                            IF #statSendBufferPos + #tempBytesUsedUtf8 <=  THEN
                              #statUserNamePos += 1;
                              CASE #tempBytesUsedUtf8 OF
                                :  // Statement section case 1
                                  #statSendBuffer[#statSendBufferPos] := #tempConvertedUtf8.%B0;
                                  #statSendBufferPos += 1;
                                :
                                  #statSendBuffer[#statSendBufferPos] := #tempConvertedUtf8.%B0;
                                  #statSendBufferPos += 1;
                                  #statSendBuffer[#statSendBufferPos] := #tempConvertedUtf8.%B1;
                                  #statSendBufferPos += 1;
                                :  // Statement section case 2 to 4
                                  #statSendBuffer[#statSendBufferPos] := #tempConvertedUtf8.%B0;
                                  #statSendBufferPos += 1;
                                  #statSendBuffer[#statSendBufferPos] := #tempConvertedUtf8.%B1;
                                  #statSendBufferPos += 1;
                                  #statSendBuffer[#statSendBufferPos] := #tempConvertedUtf8.%B2;
                                  #statSendBufferPos += 1;
                                ELSE  // Statement section ELSE
                                  ;
                              END_CASE;
                            ELSE
                              //When buffer full
                              EXIT;
                            END_IF;
                          END_FOR;
                          IF #statUserNamePos >= LEN(#username) THEN
                            #statUserNameEncodeState := ;
                          END_IF;

                        ELSE  // Statement section ELSE
                          ;
                      END_CASE;
                    END_IF;

                    // Password
                    // If the Password Flag is set to 1, the Password the next field in the payload. It must be > 0 Bytes
                    //Password field contains 0 to 65535 bytes OF binary data prefixed with a two Byte length field which indicates the number OF bytes used

                    IF #statClientIdEncodeState =
                      AND (#statWillTopicEncodeState =  OR #statWillTopicEncodeState = )
                      AND (#statWillMessageEncodeState =  OR #statWillMessageEncodeState = )
                      AND (#statUserNameEncodeState =  OR #statUserNameEncodeState = )
                      AND #statSendBufferPos <=  -  THEN
                      //When Will Topic and Will Message is encoded and buffer not full
                      CASE #statPasswordEncodeState OF
                        :  // Statement section case 1
                          //ADD len info into paket

                          #tempWordForSliceAddress := UINT_TO_WORD(#statPasswordLenUtf8Encoded);
                          #statSendBuffer[#statSendBufferPos] := #tempWordForSliceAddress.%B1; //MSB
                          #statSendBufferPos += 1;
                          #statSendBuffer[#statSendBufferPos] := #tempWordForSliceAddress.%B0; // LSB
                          #statSendBufferPos += 1;

                          FOR #tempLoopCounter := #statPasswordPos TO LEN(#password) DO
                            LMQTT_ConvertToUtf8(character     := #password[#tempLoopCounter],
                                                  convertedUtf8 => #tempConvertedUtf8,
                                                  bytesUsed     => #tempBytesUsedUtf8,
                                                  error         => #tempErrorConvertUtf8,
                                                  status        => #tempStatusConvertUtf8);

                            IF #statSendBufferPos + #tempBytesUsedUtf8 <=  THEN
                              //Increment when successful
                              #statPasswordPos += 1;

                              CASE #tempBytesUsedUtf8 OF
                                :  // Statement section case 1
                                  #statSendBuffer[#statSendBufferPos] := #tempConvertedUtf8.%B0;
                                  #statSendBufferPos += 1;
                                :
                                  #statSendBuffer[#statSendBufferPos] := #tempConvertedUtf8.%B0;
                                  #statSendBufferPos += 1;
                                  #statSendBuffer[#statSendBufferPos] := #tempConvertedUtf8.%B1;
                                  #statSendBufferPos += 1;
                                :  // Statement section case 2 to 4
                                  #statSendBuffer[#statSendBufferPos] := #tempConvertedUtf8.%B0;
                                  #statSendBufferPos += 1;
                                  #statSendBuffer[#statSendBufferPos] := #tempConvertedUtf8.%B1;
                                  #statSendBufferPos += 1;
                                  #statSendBuffer[#statSendBufferPos] := #tempConvertedUtf8.%B2;
                                  #statSendBufferPos += 1;
                                ELSE  // Statement section ELSE
                                  ;
                              END_CASE;
                            ELSE
                              //When buffer full
                              #statPasswordEncodeState := ;
                              EXIT;
                            END_IF;
                          END_FOR;

                          IF #statPasswordPos >= LEN(#password) THEN
                            #statPasswordEncodeState := ;
                          END_IF;

                        :  // Statement section case 2 to 4
                          FOR #tempLoopCounter := #statPasswordPos TO LEN(#password) DO
                            LMQTT_ConvertToUtf8(character     := #password[#tempLoopCounter],
                                                  convertedUtf8 => #tempConvertedUtf8,
                                                  bytesUsed     => #tempBytesUsedUtf8,
                                                  error         => #tempErrorConvertUtf8,
                                                  status        => #tempStatusConvertUtf8);

                            IF #statSendBufferPos + #tempBytesUsedUtf8 <=  THEN
                              #statPasswordPos += 1;
                              CASE #tempBytesUsedUtf8 OF
                                :  // Statement section case 1
                                  #statSendBuffer[#statSendBufferPos] := #tempConvertedUtf8.%B0;
                                  #statSendBufferPos += 1;
                                :
                                  #statSendBuffer[#statSendBufferPos] := #tempConvertedUtf8.%B0;
                                  #statSendBufferPos += 1;
                                  #statSendBuffer[#statSendBufferPos] := #tempConvertedUtf8.%B1;
                                  #statSendBufferPos += 1;
                                :  // Statement section case 2 to 4
                                  #statSendBuffer[#statSendBufferPos] := #tempConvertedUtf8.%B0;
                                  #statSendBufferPos += 1;
                                  #statSendBuffer[#statSendBufferPos] := #tempConvertedUtf8.%B1;
                                  #statSendBufferPos += 1;
                                  #statSendBuffer[#statSendBufferPos] := #tempConvertedUtf8.%B2;
                                  #statSendBufferPos += 1;
                                ELSE  // Statement section ELSE
                                  ;
                              END_CASE;
                            ELSE
                              //When buffer full
                              EXIT;
                            END_IF;
                          END_FOR;
                          IF #statPasswordPos >= LEN(#password) THEN
                            #statPasswordEncodeState := ;
                          END_IF;

                        ELSE  // Statement section ELSE
                          ;
                      END_CASE;
                    END_IF;

                    //set Sendlen for TSendC Block
                    #statTsendcLen := #statSendBufferPos; // Buffer pos equals amount of elements in send array
                    //reset buffer pos
                    #statSendBufferPos := 0;
                    //enable Send Req
                    #statTsendcReq := TRUE;
                    //Set Watchdog
                    #statEnableTimerCommandWatchdog := TRUE;
                    //wait for send to be done
                    #statMqttConnectState := ;
                  END_IF;
                END_REGION BUILD_CONNECT_PAKET

              :
                REGION SEND_CONNECT_PAKET_WAIT_FOR_CONNACK
                  //check tsend status
                  IF NOT #tempTsendcBusy AND #tempTsendcStatus =  THEN
                    IF (#statClientIdEncodeState =  OR #statClientIdEncodeState = )
                      AND (#statWillTopicEncodeState =  OR #statWillTopicEncodeState = )
                      AND (#statWillMessageEncodeState =  OR #statWillMessageEncodeState = )
                      AND (#statUserNameEncodeState =  OR #statUserNameEncodeState = )
                      AND (#statPasswordEncodeState =  OR #statPasswordEncodeState = ) THEN
                      //Encoding done all sent
                      #statPaketHeaderEncodeDone := FALSE;
                    ELSE
                      // More to Encode and send
                      #statEnableTimerCommandWatchdog := FALSE;
                      #statMqttConnectState := ;
                    END_IF;
                  END_IF;
                  //Check watchdog
                  IF #instTimerCommandWatchdog.Q THEN
                    #statEnableTimerCommandWatchdog := FALSE;
                    #statPaketHeaderEncodeDone := FALSE;
                    #statStatus := ; // Set correct status that identifies error clearly
                    #statSubfunctionStatus := ; // Status or return value of called FBs, FCs and system blocks
                    #statFBErrorState := #statFBState; // Set error state number for diagnostic
                    #statErrorAutoCleared := TRUE;
                    #statMqttConnectState := ;

                  END_IF;

                  //Check Connect ACK paket
                  CASE #tempMqttConnAckRcvStatus OF
                    :  //  IDLE
                      ;
                    :  // Statement section case 2 to 4
                      //disable watchdog
                      #statEnableTimerCommandWatchdog := FALSE;
                      //Encoding done all sent
                      #statPaketHeaderEncodeDone := FALSE;
                      //Go to Connected
                      #statMqttConnectState := ;
                      #statStatus := ;
                  END_CASE;
                END_REGION REGION SEND_CONNECT_PAKET

              :
                REGION CONNECTED
                  //Check Rising edge of input commands
                  #tempCommandInput.%X0 := #tempPublish AND NOT #statPublishOld;
                  #tempCommandInput.%X1 := #tempSubscribe AND NOT #statSubscribeOld;
                  #tempCommandInput.%X2 := #tempUnsubscribe AND NOT #statUnsubscribeOld;

                  //Start the keepalive timer if used
                  #statEnableMqttKeepAliveTimer := #statMqttKeepAliveUsed;

                  //set status to connected after successfully executed job
                  IF #statStatus =  THEN
                    #statStatus := ;
                  END_IF;

                  //Reset done bit
                  IF #statDone = TRUE
                    AND #tempPublish = FALSE AND #tempSubscribe = FALSE AND #tempUnsubscribe = FALSE
                  THEN
                    #statDone := FALSE;
                  END_IF;

                  REGION MQTT_COMMANDS
                    //When state machine is ready for a new input then assign correct command
                    //Ping job can be overwritten by a command.
                    IF #tempCommandInput <>
                      AND (#statMqttCommandState =  OR #statMqttCommandState = )
                    THEN
                      // New Input set, reset done flag
                      #statDone := FALSE;
                      #statMqttCommandState := BYTE_TO_DINT(#tempCommandInput);
                    END_IF;

                    CASE #statMqttCommandState OF
                      :
                        //EMPTY STATE
                        ;
                      :  // Statement section case 1
                        REGION PUBLISH_TO_TOPIC
                          //Remaining Length is the length of the variable header (TOPIC NAME + PacketID) plus the length of the Payload.
                          //Max Len of Mqtt pakets is per Standard 268,435,455 Bytes (ff,ff,ff,7f)
                          //Calculate Remain Len will be
                          //Len of TOPIC   (max 3*16382 WChars= 49.146 Bytes)
                          //plus Len of PacketID (2 Bytes)
                          //plus Len of Payload (max 268,435,455 - 49.146 - 2 = 268.386.307 Bytes ca. 268 MB)
                          //Max Array / DB Len in TIA portal is around 16 MB or 16.777.216 Byte
                          //Set Status
                          #statStatus := ;

                          // Must obey, if not currently sending PubAck Msg on a subscription
                          // Else, try in the next cycle
                          IF #tempTsendcBusy = FALSE // when tsendC is ready
                            AND #tempTsendcDone = FALSE // tsendC did not finish in this cycle
                            AND #statTsendcReq = FALSE // TsendC request was not already requested by pub ack msg
                          THEN
                            IF #statPaketHeaderEncodeDone = FALSE THEN

                              //Init
                              #statSendPaketTotalRemLen := 0;
                              #statSendBufferPos := 0;
                              #statPublishQos := #qos;
                              #statPublishMessageCnt := #publishMsgLen;
                              #statPublishTopicEncodeState := ;
                              #statPublishTopicPos := ;
                              #statPublishTopicLenUtf8Encoded := 0;
                              #statPaketId += 1;//increment
                              #statPaketIdEncoded := FALSE;
                              #statPublishEncodeMessageState := ; // No len info necessary so start directly at subsequent.
                              #statPublishMessagePos := 0; // first array element

                              //verify PayloadLen
                              #tempMaxPublishDataArrayLen := ABS(UPPER_BOUND(ARR := #publishMsgPayload, DIM := ) - LOWER_BOUND(ARR := #publishMsgPayload, DIM := )) + ;

                              //check necessary boundaries
                              IF #tempMaxPublishDataArrayLen < #statPublishMessageCnt THEN
                                #statStatus := ; // Set correct status that identifies error clearly
                                #statSubfunctionStatus := ; // Status or return value of called FBs, FCs and system blocks
                                #statFBErrorState := #statFBState; // Set error state number for diagnostic
                                #statErrorAutoCleared := TRUE;
                                #statMqttCommandState := ;
                              ELSIF LEN(#mqttTopic) =  THEN
                                #statStatus := ; // Set correct status that identifies error clearly
                                #statSubfunctionStatus := ; // Status or return value of called FBs, FCs and system blocks
                                #statFBErrorState := #statFBState; // Set error state number for diagnostic
                                #statErrorAutoCleared := TRUE;
                                #statMqttCommandState := ;
                              ELSIF #statPublishQos >  THEN
                                #statStatus := ; // Set correct status that identifies error clearly
                                #statSubfunctionStatus := ; // Status or return value of called FBs, FCs and system blocks
                                #statFBErrorState := #statFBState; // Set error state number for diagnostic
                                #statErrorAutoCleared := TRUE;
                                #statMqttCommandState := ;
                              ELSE // All ok
                                //Add amount of bytes for publish message
                                #statSendPaketTotalRemLen := #statSendPaketTotalRemLen + #statPublishMessageCnt;
                                //add publish  topic len
                                FOR #tempLoopCounter :=  TO LEN(#mqttTopic) DO
                                  LMQTT_ConvertToUtf8(character     := #mqttTopic[#tempLoopCounter],
                                                        convertedUtf8 => #tempConvertedUtf8,
                                                        bytesUsed     => #tempBytesUsedUtf8,
                                                        error         => #tempErrorConvertUtf8,
                                                        status        => #tempStatusConvertUtf8);
                                  #statPublishTopicLenUtf8Encoded := #statPublishTopicLenUtf8Encoded + #tempBytesUsedUtf8;
                                END_FOR;
                                #statSendPaketTotalRemLen := #statSendPaketTotalRemLen + #statPublishTopicLenUtf8Encoded + ;

                                //Build Publish Telegram
                                //Fixed Header - Write Paket Type
                                #statSendBuffer[#statSendBufferPos] := ;
                                // Set DUP flag always to FALSE
                                #statSendBuffer[#statSendBufferPos].%X3 := FALSE;
                                // Set QoS Level
                                CASE #statPublishQos OF
                                  :  // Statement section case 0
                                    #statSendBuffer[#statSendBufferPos].%X2 := FALSE;
                                    #statSendBuffer[#statSendBufferPos].%X1 := FALSE;
                                  :  // Statement section case 1
                                    #statSendBuffer[#statSendBufferPos].%X2 := FALSE;
                                    #statSendBuffer[#statSendBufferPos].%X1 := TRUE;
                                    //Add two byte len info for Mandatory packet ID
                                    #statSendPaketTotalRemLen := #statSendPaketTotalRemLen + ;
                                  : // Statement section case 2
                                    #statSendBuffer[#statSendBufferPos].%X2 := TRUE;
                                    #statSendBuffer[#statSendBufferPos].%X1 := FALSE;
                                    //Add two byte len info for Mandatory packet ID
                                    #statSendPaketTotalRemLen := #statSendPaketTotalRemLen + ;
                                  ELSE
                                    ;
                                END_CASE;
                                //Set retain bit
                                #statSendBuffer[#statSendBufferPos].%X0 := #retain;

                                #statSendBufferPos += 1; // increment

                                //Write Remaining Paket Len info
                                WHILE (#statSendPaketTotalRemLen > )
                                DO//See MQTT Spec for explanation of this calculation
                                  #statEncodedRemPaketLenAsByte := UDINT_TO_BYTE(#statSendPaketTotalRemLen MOD );
                                  #statSendPaketTotalRemLen := #statSendPaketTotalRemLen / ;
                                  // if there are more data to encode, set the top bit of this byte
                                  IF #statSendPaketTotalRemLen >
                                  THEN
                                    // Do this and continue while loop
                                    #statEncodedRemPaketLenAsByte := #statEncodedRemPaketLenAsByte OR UDINT_TO_BYTE();
                                    #statSendBuffer[#statSendBufferPos] := #statEncodedRemPaketLenAsByte;
                                    #statSendBufferPos += 1;
                                  ELSE
                                    //do this and leave while loop
                                    #statSendBuffer[#statSendBufferPos] := #statEncodedRemPaketLenAsByte;
                                    #statSendBufferPos += 1;
                                  END_IF;
                                END_WHILE;
                                //When all done, set encode to true
                                #statPaketHeaderEncodeDone := TRUE;
                              END_IF;
                            END_IF;

                            //Header Encoded - now Topic, PacketId and Message need to be encoded.
                            IF #statPaketHeaderEncodeDone = TRUE THEN

                              //Publish Topic
                              IF #statSendBufferPos <=  -  THEN
                                CASE #statPublishTopicEncodeState OF
                                  :  // Statement section case 1
                                    //ADD len info into paket

                                    #tempWordForSliceAddress := UINT_TO_WORD(#statPublishTopicLenUtf8Encoded);
                                    #statSendBuffer[#statSendBufferPos] := #tempWordForSliceAddress.%B1; //MSB
                                    #statSendBufferPos += 1;
                                    #statSendBuffer[#statSendBufferPos] := #tempWordForSliceAddress.%B0; // LSB
                                    #statSendBufferPos += 1;

                                    FOR #tempLoopCounter := #statPublishTopicPos TO LEN(#mqttTopic) DO
                                      LMQTT_ConvertToUtf8(character     := #mqttTopic[#tempLoopCounter],
                                                            convertedUtf8 => #tempConvertedUtf8,
                                                            bytesUsed     => #tempBytesUsedUtf8,
                                                            error         => #tempErrorConvertUtf8,
                                                            status        => #tempStatusConvertUtf8);

                                      IF #statSendBufferPos + #tempBytesUsedUtf8 <=  THEN
                                        #statPublishTopicPos += 1;
                                        CASE #tempBytesUsedUtf8 OF
                                          :  // Statement section case 1
                                            #statSendBuffer[#statSendBufferPos] := #tempConvertedUtf8.%B0;
                                            #statSendBufferPos += 1;
                                          :
                                            #statSendBuffer[#statSendBufferPos] := #tempConvertedUtf8.%B0;
                                            #statSendBufferPos += 1;
                                            #statSendBuffer[#statSendBufferPos] := #tempConvertedUtf8.%B1;
                                            #statSendBufferPos += 1;
                                          :  // Statement section case 2 to 4
                                            #statSendBuffer[#statSendBufferPos] := #tempConvertedUtf8.%B0;
                                            #statSendBufferPos += 1;
                                            #statSendBuffer[#statSendBufferPos] := #tempConvertedUtf8.%B1;
                                            #statSendBufferPos += 1;
                                            #statSendBuffer[#statSendBufferPos] := #tempConvertedUtf8.%B2;
                                            #statSendBufferPos += 1;
                                          ELSE  // Statement section ELSE
                                            ;
                                        END_CASE;
                                      ELSE
                                        //When buffer full
                                        #statPublishTopicEncodeState := ;
                                        EXIT;
                                      END_IF;
                                    END_FOR;
                                    IF #statPublishTopicPos >= LEN(#mqttTopic) THEN
                                      #statPublishTopicEncodeState := ;
                                    END_IF;


                                  :  // Statement section case 2 to 4
                                    FOR #tempLoopCounter := #statPublishTopicPos TO LEN(#mqttTopic) DO

                                      LMQTT_ConvertToUtf8(character     := #mqttTopic[#tempLoopCounter],
                                                            convertedUtf8 => #tempConvertedUtf8,
                                                            bytesUsed     => #tempBytesUsedUtf8,
                                                            error         => #tempErrorConvertUtf8,
                                                            status        => #tempStatusConvertUtf8);
                                      IF #statSendBufferPos + #tempBytesUsedUtf8 <=  THEN
                                        #statPublishTopicPos += 1;
                                        CASE #tempBytesUsedUtf8 OF
                                          :  // Statement section case 1
                                            #statSendBuffer[#statSendBufferPos] := #tempConvertedUtf8.%B0;
                                            #statSendBufferPos += 1;
                                          :
                                            #statSendBuffer[#statSendBufferPos] := #tempConvertedUtf8.%B0;
                                            #statSendBufferPos += 1;
                                            #statSendBuffer[#statSendBufferPos] := #tempConvertedUtf8.%B1;
                                            #statSendBufferPos += 1;
                                          :  // Statement section case 2 to 4
                                            #statSendBuffer[#statSendBufferPos] := #tempConvertedUtf8.%B0;
                                            #statSendBufferPos += 1;
                                            #statSendBuffer[#statSendBufferPos] := #tempConvertedUtf8.%B1;
                                            #statSendBufferPos += 1;
                                            #statSendBuffer[#statSendBufferPos] := #tempConvertedUtf8.%B2;
                                            #statSendBufferPos += 1;
                                          ELSE  // Statement section ELSE
                                            ;
                                        END_CASE;
                                      ELSE
                                        //When buffer full
                                        EXIT;
                                      END_IF;
                                    END_FOR;
                                    IF #statPublishTopicPos >= LEN(#mqttTopic) THEN
                                      #statPublishTopicEncodeState := ;
                                    END_IF;
                                  ELSE  // SKIP if done
                                    ;
                                END_CASE;
                              END_IF;

                              // Encode MessageID, when QOS > 0 and  Topic done and buffer not full
                              IF #statPublishTopicEncodeState =
                                AND #statPaketIdEncoded = FALSE
                                AND #statSendBufferPos <=  -  THEN
                                // Check QoS - only necessary if QoS >0
                                CASE #statPublishQos OF
                                  :
                                    #tempWordForSliceAddress := UINT_TO_WORD(#statPaketId);
                                    #statSendBuffer[#statSendBufferPos] := #tempWordForSliceAddress.%B1; //MSB
                                    #statSendBufferPos += 1;
                                    #statSendBuffer[#statSendBufferPos] := #tempWordForSliceAddress.%B0; //LSB
                                    #statSendBufferPos += 1;
                                  :
                                    #tempWordForSliceAddress := UINT_TO_WORD(#statPaketId);
                                    #statSendBuffer[#statSendBufferPos] := #tempWordForSliceAddress.%B1; //MSB
                                    #statSendBufferPos += 1;
                                    #statSendBuffer[#statSendBufferPos] := #tempWordForSliceAddress.%B0; //LSB
                                    #statSendBufferPos += 1;
                                  ELSE
                                    //No paket id to encode here
                                    ;
                                END_CASE;
                                //Finally:
                                #statPaketIdEncoded := TRUE;
                              END_IF;

                              // Encode Payload, when  Topic done and PaketID Done and buffer not full
                              IF #statPublishTopicEncodeState =
                                AND #statPaketIdEncoded = TRUE
                                AND #statSendBufferPos <  THEN

                                // Publish Message Encoding
                                // This Contains the payload from the publish message expressed as a sequence bytes.
                                CASE #statPublishEncodeMessageState OF
                                  :  // Statement section case 2 to 4
                                    #tempLowerBoundPublishDataArray := LOWER_BOUND(ARR := #publishMsgPayload, DIM := );

                                    FOR #tempLoopCounter := #statPublishMessagePos TO UDINT_TO_DINT(#statPublishMessageCnt - 1) DO
                                      IF #statSendBufferPos <=  THEN
                                        #statSendBuffer[#statSendBufferPos] := #publishMsgPayload[#tempLowerBoundPublishDataArray + #tempLoopCounter];
                                        #statSendBufferPos += 1;
                                        //Increment when successful
                                        #statPublishMessagePos += 1;
                                      ELSE
                                        //When Buffer Full
                                        EXIT;
                                      END_IF;
                                    END_FOR;
                                    // If everything was copied successfull
                                    IF #statPublishMessagePos >= #statPublishMessageCnt THEN
                                      #statPublishEncodeMessageState := ;
                                    END_IF;
                                  ELSE  // Statement section ELSE
                                    ;
                                END_CASE;
                              END_IF;

                              //set Sendlen for TSendC Block
                              #statTsendcLen := #statSendBufferPos; // Buffer pos equals amount of elements in send array
                              //reset buffer pos
                              #statSendBufferPos := 0;
                              //enable Send Req
                              #statTsendcReq := TRUE;
                              //Set Watchdog
                              #statEnableTimerCommandWatchdog := TRUE;
                              //wait for send to be done
                              #statMqttCommandState := ;
                            END_IF;
                          END_IF;
                        END_REGION PUBLISH_TO_TOPIC

                      :
                        REGION SEND_PUBLISH_WAIT_FOR_RESPONSE
                          //check tsend status
                          IF NOT #tempTsendcBusy AND #tempTsendcStatus =  THEN

                            IF (#statPublishTopicEncodeState = )
                              AND (#statPublishEncodeMessageState = ) THEN
                              //Encoding done all sent
                              #statPaketHeaderEncodeDone := FALSE;
                              //  with QoS = 0 Job done
                              IF #statPublishQos =  THEN
                                // job done
                                #statDone := TRUE;
                                // go back to idle
                                #statMqttCommandState := ;
                                //reset Watchdog
                                #statEnableTimerCommandWatchdog := FALSE;
                                // Set Status back to connected
                                #statStatus := ;
                              END_IF;
                            ELSE
                              // More to Encode and send
                              #statEnableTimerCommandWatchdog := FALSE;
                              #statMqttCommandState := ;
                            END_IF;

                          END_IF;
                          IF (#instTsendC.STATUS =  OR #instTsendC.STATUS =)THEN
                            #statPubRecReady := 1;
                          ELSE
                            #statPubRecReady := 0;

                          END_IF;

                          //check watchdog
                          IF #instTimerCommandWatchdog.Q THEN
                            #statEnableTimerCommandWatchdog := FALSE;
                            #statStatus := ; // Set correct status that identifies error clearly
                            #statSubfunctionStatus := ; // Status or return value of called FBs, FCs and system blocks
                            #statFBErrorState := #statFBState; // Set error state number for diagnostic
                            #statErrorAutoCleared := TRUE;
                            #statMqttCommandState := ;


                          END_IF;

                          //When QoS = 1; Wait for Publish ACK paket
                          CASE #tempMqttPubAckRcv OF
                            :  // Statement section case 0 IDLE
                              ;
                            :  // Statement section case 1 OKAY
                              //disable watchdog
                              #statEnableTimerCommandWatchdog := FALSE;
                              //Encoding done all sent
                              #statPaketHeaderEncodeDone := FALSE;
                              //Publish QoS 1 = Done
                              #statDone := TRUE;
                              #statMqttCommandState := ;
                              // Set Status back to connected
                              #statStatus := ;
                            :
                              #statStatus := ; // Set correct status that identifies error clearly
                              #statSubfunctionStatus := ; // Status or return value of called FBs, FCs and system blocks
                              #statFBErrorState := #statFBState; // Set error state number for diagnostic
                              #statErrorAutoCleared := TRUE;
                              #statMqttCommandState := ;
                          END_CASE;

                          //When QOS = 2 and Pub Rec Receieved:
                          CASE #statMqttPubRecRcv OF
                            :  // 0 IDLE
                              ;
                            :
                              IF (#statPubRecReady) THEN
                                //Encoding done all sent
                                #statPaketHeaderEncodeDone := FALSE;
                                // Send Publish Release paket
                                #statSendBufferPos := 0;
                                #statSendBuffer[#statSendBufferPos] := ;
                                #statSendBufferPos += 1;
                                //Remaining Lenght (must be 2)
                                #statSendBuffer[#statSendBufferPos] := ;
                                #statSendBufferPos += 1;
                                // add paket id
                                #tempWordForSliceAddress := UINT_TO_WORD(#statPaketId);
                                #statSendBuffer[#statSendBufferPos] := #tempWordForSliceAddress.%B1; //MSB
                                #statSendBufferPos += 1;
                                #statSendBuffer[#statSendBufferPos] := #tempWordForSliceAddress.%B0; //LSB
                                #statSendBufferPos += 1;
                                #statTsendcLen := #statSendBufferPos;
                                //Start send request
                                #statTsendcReq := TRUE;
                                #statMqttPubRecRcv := 0;
                                #statPubRecReady := 0;




                                //Reset watchdog and start
                                RESET_TIMER(#instTimerCommandWatchdog);
                                #statEnableTimerCommandWatchdog := TRUE;
                              END_IF;
                              //Stay in State
                            :
                              #statStatus := ; // Set correct status that identifies error clearly
                              #statSubfunctionStatus := ; // Status or return value of called FBs, FCs and system blocks
                              #statFBErrorState := #statFBState; // Set error state number for diagnostic
                              #statErrorAutoCleared := TRUE;
                              #statMqttCommandState := ;
                          END_CASE;

                          //When QOS = 2 and Pub Complete Receieved:
                          CASE #tempMqttPubCompRcv OF
                            :  // Idle
                              ;
                            :  //When QOS = 2 and Pub Complete Receieved:
                              //disable watchdog
                              #statEnableTimerCommandWatchdog := FALSE;
                              //Encoding done all sent
                              #statPaketHeaderEncodeDone := FALSE;
                              //Publish QoS 2 = Done
                              #statDone := TRUE;

                              #statMqttCommandState := ;
                              // Set Status back to connected
                              #statStatus := ;
                            :
                              #statStatus := ; // Set correct status that identifies error clearly
                              #statSubfunctionStatus := ; // Status or return value of called FBs, FCs and system blocks
                              #statFBErrorState := #statFBState; // Set error state number for diagnostic
                              #statErrorAutoCleared := TRUE;
                              #statMqttCommandState := ;
                          END_CASE;
                        END_REGION MQTT_COMMAND_SEND_PUBLISH

                      :  // Statement section case 2
                        REGION SUBSCRIBE_TO_TOPIC
                          //Remaining Length is the length of the variable header (PacketID, 2Bytes) plus the length of the Payload.
                          //Max Len of Mqtt pakets is per Standard 268,435,455 Bytes (ff,ff,ff,7f)
                          //Calculate Remain Len will be
                          //Len of TOPIC   (max 3*16382 WChars= 49.146 Bytes)
                          //LenInfo Topic (2Byte)
                          //QoS of Topic (1Byte)
                          //
                          //Set Status
                          #statStatus := ;
                          // Must obey, if not currently sending PubAck Msg on a subscription
                          // Else, try in the next cycle
                          IF #tempTsendcBusy = FALSE // when tsendC is ready
                            AND #tempTsendcDone = FALSE // tsendC did not finish in this cycle
                            AND #statTsendcReq = FALSE // TsendC request was not already requested by pub ack msg
                          THEN
                            IF #statPaketHeaderEncodeDone = FALSE THEN

                              //Init
                              #statSendPaketTotalRemLen := 0;
                              #statSendBufferPos := 0;
                              #statSubscribeQos := #qos;
                              #statSubscribeTopicEncodeState := ;
                              #statSubscribeTopicPos := ;
                              #statSubscribeTopicLenUtf8Encoded := 0;
                              #statPaketId += 1;//increment
                              #statSubscribeQosEncoded := FALSE;

                              //check necessary boundaries

                              IF LEN(#mqttTopic) =  THEN
                                #statStatus := ; // Set correct status that identifies error clearly
                                #statSubfunctionStatus := ; // Status or return value of called FBs, FCs and system blocks
                                #statFBErrorState := #statFBState; // Set error state number for diagnostic
                                #statErrorAutoCleared := TRUE;
                                #statMqttCommandState := ;
                              ELSIF #statSubscribeQos >  THEN
                                #statStatus := ; // Set correct status that identifies error clearly
                                #statSubfunctionStatus := ; // Status or return value of called FBs, FCs and system blocks
                                #statFBErrorState := #statFBState; // Set error state number for diagnostic
                                #statErrorAutoCleared := TRUE;
                                #statMqttCommandState := ;
                              ELSE // All ok
                                //Add two Byte for Paket ID:
                                #statSendPaketTotalRemLen := #statSendPaketTotalRemLen + ;
                                //Add one Byte for QoS Info:
                                #statSendPaketTotalRemLen := #statSendPaketTotalRemLen + ;
                                //add subscribe  topic len
                                FOR #tempLoopCounter :=  TO LEN(#mqttTopic) DO
                                  LMQTT_ConvertToUtf8(character     := #mqttTopic[#tempLoopCounter],
                                                        convertedUtf8 => #tempConvertedUtf8,
                                                        bytesUsed     => #tempBytesUsedUtf8,
                                                        error         => #tempErrorConvertUtf8,
                                                        status        => #tempStatusConvertUtf8);
                                  #statSubscribeTopicLenUtf8Encoded := #statSubscribeTopicLenUtf8Encoded + #tempBytesUsedUtf8;
                                END_FOR;
                                //Add len of topic plus len info
                                #statSendPaketTotalRemLen := #statSendPaketTotalRemLen + #statSubscribeTopicLenUtf8Encoded + ;

                                //Build Subscribe Telegram
                                //Fixed Header - Write Paket Type
                                #statSendBuffer[#statSendBufferPos] := ;
                                #statSendBufferPos += 1; // increment

                                //Write Remaining Paket Len info
                                WHILE (#statSendPaketTotalRemLen > )
                                DO//See MQTT Spec for explanation of this calculation
                                  #statEncodedRemPaketLenAsByte := UDINT_TO_BYTE(#statSendPaketTotalRemLen MOD );
                                  #statSendPaketTotalRemLen := #statSendPaketTotalRemLen / ;
                                  // if there are more data to encode, set the top bit of this byte
                                  IF #statSendPaketTotalRemLen >
                                  THEN
                                    // Do this and continue while loop
                                    #statEncodedRemPaketLenAsByte := #statEncodedRemPaketLenAsByte OR UDINT_TO_BYTE();
                                    #statSendBuffer[#statSendBufferPos] := #statEncodedRemPaketLenAsByte;
                                    #statSendBufferPos += 1;
                                  ELSE
                                    //do this and leave while loop
                                    #statSendBuffer[#statSendBufferPos] := #statEncodedRemPaketLenAsByte;
                                    #statSendBufferPos += 1;
                                  END_IF;
                                END_WHILE;

                                // Set Paket Id
                                #tempWordForSliceAddress := UINT_TO_WORD(#statPaketId);
                                #statSendBuffer[#statSendBufferPos] := #tempWordForSliceAddress.%B1; //MSB
                                #statSendBufferPos += 1;
                                #statSendBuffer[#statSendBufferPos] := #tempWordForSliceAddress.%B0; //LSB
                                #statSendBufferPos += 1;

                                //When all done, set encode to true
                                #statPaketHeaderEncodeDone := TRUE;
                              END_IF;
                            END_IF;
                            //Header Encoded
                            IF #statPaketHeaderEncodeDone = TRUE THEN
                              //Header Encoded - now Topic and qos encoding

                              //Subscribe Topic
                              IF #statSendBufferPos <=  -  THEN
                                CASE #statSubscribeTopicEncodeState OF
                                  :  // Statement section case 1
                                    //ADD len info into paket

                                    #tempWordForSliceAddress := UINT_TO_WORD(#statSubscribeTopicLenUtf8Encoded);
                                    #statSendBuffer[#statSendBufferPos] := #tempWordForSliceAddress.%B1; //MSB
                                    #statSendBufferPos += 1;
                                    #statSendBuffer[#statSendBufferPos] := #tempWordForSliceAddress.%B0; // LSB
                                    #statSendBufferPos += 1;

                                    FOR #tempLoopCounter := #statSubscribeTopicPos TO LEN(#mqttTopic) DO
                                      LMQTT_ConvertToUtf8(character     := #mqttTopic[#tempLoopCounter],
                                                            convertedUtf8 => #tempConvertedUtf8,
                                                            bytesUsed     => #tempBytesUsedUtf8,
                                                            error         => #tempErrorConvertUtf8,
                                                            status        => #tempStatusConvertUtf8);

                                      IF #statSendBufferPos + #tempBytesUsedUtf8 <=  THEN
                                        #statSubscribeTopicPos += 1;
                                        CASE #tempBytesUsedUtf8 OF
                                          :  // Statement section case 1
                                            #statSendBuffer[#statSendBufferPos] := #tempConvertedUtf8.%B0;
                                            #statSendBufferPos += 1;
                                          :
                                            #statSendBuffer[#statSendBufferPos] := #tempConvertedUtf8.%B0;
                                            #statSendBufferPos += 1;
                                            #statSendBuffer[#statSendBufferPos] := #tempConvertedUtf8.%B1;
                                            #statSendBufferPos += 1;
                                          :  // Statement section case 2 to 4
                                            #statSendBuffer[#statSendBufferPos] := #tempConvertedUtf8.%B0;
                                            #statSendBufferPos += 1;
                                            #statSendBuffer[#statSendBufferPos] := #tempConvertedUtf8.%B1;
                                            #statSendBufferPos += 1;
                                            #statSendBuffer[#statSendBufferPos] := #tempConvertedUtf8.%B2;
                                            #statSendBufferPos += 1;
                                          ELSE  // Statement section ELSE
                                            ;
                                        END_CASE;
                                      ELSE
                                        //When buffer full
                                        #statSubscribeTopicEncodeState := ;
                                        EXIT;
                                      END_IF;
                                    END_FOR;
                                    IF #statSubscribeTopicPos >= LEN(#mqttTopic) THEN
                                      #statSubscribeTopicEncodeState := ;
                                    END_IF;

                                  :  // Statement section case 2 to 4
                                    FOR #tempLoopCounter := #statSubscribeTopicPos TO LEN(#mqttTopic) DO

                                      LMQTT_ConvertToUtf8(character     := #mqttTopic[#tempLoopCounter],
                                                            convertedUtf8 => #tempConvertedUtf8,
                                                            bytesUsed     => #tempBytesUsedUtf8,
                                                            error         => #tempErrorConvertUtf8,
                                                            status        => #tempStatusConvertUtf8);
                                      IF #statSendBufferPos + #tempBytesUsedUtf8 <=  THEN
                                        #statSubscribeTopicPos += 1;
                                        CASE #tempBytesUsedUtf8 OF
                                          :  // Statement section case 1
                                            #statSendBuffer[#statSendBufferPos] := #tempConvertedUtf8.%B0;
                                            #statSendBufferPos += 1;
                                          :
                                            #statSendBuffer[#statSendBufferPos] := #tempConvertedUtf8.%B0;
                                            #statSendBufferPos += 1;
                                            #statSendBuffer[#statSendBufferPos] := #tempConvertedUtf8.%B1;
                                            #statSendBufferPos += 1;
                                          :  // Statement section case 2 to 4
                                            #statSendBuffer[#statSendBufferPos] := #tempConvertedUtf8.%B0;
                                            #statSendBufferPos += 1;
                                            #statSendBuffer[#statSendBufferPos] := #tempConvertedUtf8.%B1;
                                            #statSendBufferPos += 1;
                                            #statSendBuffer[#statSendBufferPos] := #tempConvertedUtf8.%B2;
                                            #statSendBufferPos += 1;
                                          ELSE  // Statement section ELSE
                                            ;
                                        END_CASE;
                                      ELSE
                                        //When buffer full
                                        EXIT;
                                      END_IF;
                                    END_FOR;
                                    IF #statSubscribeTopicPos >= LEN(#mqttTopic) THEN
                                      #statSubscribeTopicEncodeState := ;
                                    END_IF;
                                  ELSE  // Skip when Done
                                    ;
                                END_CASE;
                              END_IF;

                              IF #statSubscribeTopicEncodeState =
                                AND #statSendBufferPos <=  -  THEN
                                #statSendBuffer[#statSendBufferPos] := USINT_TO_BYTE(#statSubscribeQos);
                                #statSendBufferPos += 1;
                                #statSubscribeQosEncoded := TRUE;
                              END_IF;


                              //set Sendlen for TSendC Block
                              #statTsendcLen := #statSendBufferPos; // Buffer pos equals amount of elements in send array
                              //reset buffer pos
                              #statSendBufferPos := 0;
                              //enable Send Req
                              #statTsendcReq := TRUE;
                              //Set Watchdog
                              #statEnableTimerCommandWatchdog := TRUE;
                              //wait for send to be done
                              #statMqttCommandState := ;
                            END_IF;
                          END_IF;
                        END_REGION SUBSCRIBE_TO_TOPIC

                      :
                        REGION SEND_SUBSCRIBE_WAIT_FOR_RESPONSE
                          //check tsend status
                          IF NOT #tempTsendcBusy AND #tempTsendcStatus =  THEN
                            IF #statSubscribeTopicEncodeState =
                              AND #statSubscribeQosEncoded = TRUE THEN
                              //Encoding done all sent
                              #statPaketHeaderEncodeDone := FALSE;
                            ELSE
                              // More to Encode and send
                              #statEnableTimerCommandWatchdog := FALSE; // reset watchdog
                              #statMqttCommandState := ;
                            END_IF;
                          END_IF;
                          //Wait for timeout
                          IF #instTimerCommandWatchdog.Q THEN
                            #statEnableTimerCommandWatchdog := FALSE;
                            #statStatus := ; // Set correct status that identifies error clearly
                            #statSubfunctionStatus := ; // Status or return value of called FBs, FCs and system blocks
                            #statFBErrorState := #statFBState; // Set error state number for diagnostic
                            #statErrorAutoCleared := TRUE;
                            #statMqttCommandState := ;
                          END_IF;

                          //Check Subscribe ACK paket
                          CASE #tempMqttSubAckRcv OF
                            :  // Statement section case 1
                              ;
                            :  // Statement section case 2 to 4
                              //disable watchdog
                              #statEnableTimerCommandWatchdog := FALSE;
                              //Encoding done all sent
                              #statPaketHeaderEncodeDone := FALSE;
                              // Job done
                              #statDone := TRUE;
                              #statMqttCommandState := ;
                              // Set Status back to connected
                              #statStatus := ;
                            :  // PaketId Invalid
                              #statStatus := ; // Set correct status that identifies error clearly
                              #statSubfunctionStatus := ; // Status or return value of called FBs, FCs and system blocks
                              #statFBErrorState := #statFBState; // Set error state number for diagnostic
                              #statErrorAutoCleared := TRUE;
                              #statMqttCommandState := ;
                            :
                              #statStatus := ; // Set correct status that identifies error clearly
                              #statSubfunctionStatus := ; // Status or return value of called FBs, FCs and system blocks
                              #statFBErrorState := #statFBState; // Set error state number for diagnostic
                              #statErrorAutoCleared := TRUE;
                              #statMqttCommandState := ;
                          END_CASE;
                        END_REGION SEND_SUBSCRIBE_WAIT_FOR_RESPONSE

                      :// Unsubscribe from topics
                        REGION UNSUBSCRIBE_FROM_TOPIC
                          //Remaining Length is the length of the variable header (PacketID, 2Bytes) plus the length of the Payload.
                          //Max Len of Mqtt pakets is per Standard 268,435,455 Bytes (ff,ff,ff,7f)
                          //Calculate Remain Len will be
                          //Len of TOPIC   (max 3*16382 WChars= 49.146 Bytes)
                          //LenInfo Topic (2Byte)
                          //
                          //Set Status
                          #statStatus := ;
                          // Must obey, if not currently sending PubAck Msg on a subscription
                          // Else, try in the next cycle
                          IF #tempTsendcBusy = FALSE // when tsendC is ready
                            AND #tempTsendcDone = FALSE // tsendC did not finish in this cycle
                            AND #statTsendcReq = FALSE // TsendC request was not already requested by pub ack msg
                          THEN
                            //Header not encoded
                            IF #statPaketHeaderEncodeDone = FALSE THEN
                              //Init
                              #statSendPaketTotalRemLen := 0;
                              #statSendBufferPos := 0;
                              #statUnsubscribeTopicEncodeState := ;
                              #statUnsubscribeTopicPos := ;
                              #statUnsubscribeTopicLenUtf8Encoded := 0;
                              #statPaketId += 1;//increment

                              //check necessary boundaries

                              IF LEN(#mqttTopic) =  THEN
                                #statStatus := ; // Set correct status that identifies error clearly
                                #statSubfunctionStatus := ; // Status or return value of called FBs, FCs and system blocks
                                #statFBErrorState := #statFBState; // Set error state number for diagnostic
                                #statErrorUserCleared := TRUE;
                              ELSE // All ok
                                //Add two Byte for Paket ID:
                                #statSendPaketTotalRemLen := #statSendPaketTotalRemLen + ;
                                //add unsubscribe  topic len
                                FOR #tempLoopCounter :=  TO LEN(#mqttTopic) DO
                                  LMQTT_ConvertToUtf8(character     := #mqttTopic[#tempLoopCounter],
                                                        convertedUtf8 => #tempConvertedUtf8,
                                                        bytesUsed     => #tempBytesUsedUtf8,
                                                        error         => #tempErrorConvertUtf8,
                                                        status        => #tempStatusConvertUtf8);
                                  #statUnsubscribeTopicLenUtf8Encoded := #statUnsubscribeTopicLenUtf8Encoded + #tempBytesUsedUtf8;
                                END_FOR;
                                //Add len of topic plus len info
                                #statSendPaketTotalRemLen := #statSendPaketTotalRemLen + #statUnsubscribeTopicLenUtf8Encoded + ;

                                //Build Subscribe Telegram
                                //Fixed Header - Write Paket Type
                                #statSendBuffer[#statSendBufferPos] := ;
                                #statSendBufferPos += 1; // increment

                                //Write Remaining Paket Len info
                                WHILE (#statSendPaketTotalRemLen > )
                                DO//See MQTT Spec for explanation of this calculation
                                  #statEncodedRemPaketLenAsByte := UDINT_TO_BYTE(#statSendPaketTotalRemLen MOD );
                                  #statSendPaketTotalRemLen := #statSendPaketTotalRemLen / ;
                                  // if there are more data to encode, set the top bit of this byte
                                  IF #statSendPaketTotalRemLen >
                                  THEN
                                    // Do this and continue while loop
                                    #statEncodedRemPaketLenAsByte := #statEncodedRemPaketLenAsByte OR UDINT_TO_BYTE();
                                    #statSendBuffer[#statSendBufferPos] := #statEncodedRemPaketLenAsByte;
                                    #statSendBufferPos += 1;
                                  ELSE
                                    //do this and leave while loop
                                    #statSendBuffer[#statSendBufferPos] := #statEncodedRemPaketLenAsByte;
                                    #statSendBufferPos += 1;
                                  END_IF;
                                END_WHILE;

                                // Set Paket Id
                                #tempWordForSliceAddress := UINT_TO_WORD(#statPaketId);
                                #statSendBuffer[#statSendBufferPos] := #tempWordForSliceAddress.%B1; //MSB
                                #statSendBufferPos += 1;
                                #statSendBuffer[#statSendBufferPos] := #tempWordForSliceAddress.%B0; //LSB
                                #statSendBufferPos += 1;

                                //When all done, set encode to true
                                #statPaketHeaderEncodeDone := TRUE;
                              END_IF;
                            END_IF;

                            //Header Encoded -
                            IF #statPaketHeaderEncodeDone = TRUE THEN
                              //Unsubscribe Topic
                              IF #statSendBufferPos <=  -  THEN
                                CASE #statUnsubscribeTopicEncodeState OF
                                  :  // Statement section case 1
                                    //ADD len info into paket

                                    #tempWordForSliceAddress := UINT_TO_WORD(#statUnsubscribeTopicLenUtf8Encoded);
                                    #statSendBuffer[#statSendBufferPos] := #tempWordForSliceAddress.%B1; //MSB
                                    #statSendBufferPos += 1;
                                    #statSendBuffer[#statSendBufferPos] := #tempWordForSliceAddress.%B0; // LSB
                                    #statSendBufferPos += 1;

                                    FOR #tempLoopCounter := #statUnsubscribeTopicPos TO LEN(#mqttTopic) DO
                                      LMQTT_ConvertToUtf8(character     := #mqttTopic[#tempLoopCounter],
                                                            convertedUtf8 => #tempConvertedUtf8,
                                                            bytesUsed     => #tempBytesUsedUtf8,
                                                            error         => #tempErrorConvertUtf8,
                                                            status        => #tempStatusConvertUtf8);

                                      IF #statSendBufferPos + #tempBytesUsedUtf8 <=  THEN
                                        #statUnsubscribeTopicPos += 1;
                                        CASE #tempBytesUsedUtf8 OF
                                          :  // Statement section case 1
                                            #statSendBuffer[#statSendBufferPos] := #tempConvertedUtf8.%B0;
                                            #statSendBufferPos += 1;
                                          :
                                            #statSendBuffer[#statSendBufferPos] := #tempConvertedUtf8.%B0;
                                            #statSendBufferPos += 1;
                                            #statSendBuffer[#statSendBufferPos] := #tempConvertedUtf8.%B1;
                                            #statSendBufferPos += 1;
                                          :  // Statement section case 2 to 4
                                            #statSendBuffer[#statSendBufferPos] := #tempConvertedUtf8.%B0;
                                            #statSendBufferPos += 1;
                                            #statSendBuffer[#statSendBufferPos] := #tempConvertedUtf8.%B1;
                                            #statSendBufferPos += 1;
                                            #statSendBuffer[#statSendBufferPos] := #tempConvertedUtf8.%B2;
                                            #statSendBufferPos += 1;
                                          ELSE  // Statement section ELSE
                                            ;
                                        END_CASE;
                                      ELSE
                                        //When buffer full
                                        #statUnsubscribeTopicEncodeState := ;
                                        EXIT;
                                      END_IF;
                                    END_FOR;
                                    IF #statUnsubscribeTopicPos >= LEN(#mqttTopic) THEN
                                      #statUnsubscribeTopicEncodeState := ;
                                    END_IF;

                                  :  // Statement section case 2 to 4
                                    FOR #tempLoopCounter := #statUnsubscribeTopicPos TO LEN(#mqttTopic) DO

                                      LMQTT_ConvertToUtf8(character     := #mqttTopic[#tempLoopCounter],
                                                            convertedUtf8 => #tempConvertedUtf8,
                                                            bytesUsed     => #tempBytesUsedUtf8,
                                                            error         => #tempErrorConvertUtf8,
                                                            status        => #tempStatusConvertUtf8);
                                      IF #statSendBufferPos + #tempBytesUsedUtf8 <=  THEN
                                        #statUnsubscribeTopicPos += 1;
                                        CASE #tempBytesUsedUtf8 OF
                                          :  // Statement section case 1
                                            #statSendBuffer[#statSendBufferPos] := #tempConvertedUtf8.%B0;
                                            #statSendBufferPos += 1;
                                          :
                                            #statSendBuffer[#statSendBufferPos] := #tempConvertedUtf8.%B0;
                                            #statSendBufferPos += 1;
                                            #statSendBuffer[#statSendBufferPos] := #tempConvertedUtf8.%B1;
                                            #statSendBufferPos += 1;
                                          :  // Statement section case 2 to 4
                                            #statSendBuffer[#statSendBufferPos] := #tempConvertedUtf8.%B0;
                                            #statSendBufferPos += 1;
                                            #statSendBuffer[#statSendBufferPos] := #tempConvertedUtf8.%B1;
                                            #statSendBufferPos += 1;
                                            #statSendBuffer[#statSendBufferPos] := #tempConvertedUtf8.%B2;
                                            #statSendBufferPos += 1;
                                          ELSE  // Statement section ELSE
                                            ;
                                        END_CASE;
                                      ELSE
                                        //When buffer full
                                        EXIT;
                                      END_IF;
                                    END_FOR;
                                    IF #statUnsubscribeTopicPos >= LEN(#mqttTopic) THEN
                                      #statUnsubscribeTopicEncodeState := ;
                                    END_IF;
                                  ELSE  // Skip when Done
                                    ;
                                END_CASE;
                              END_IF;

                              //set Sendlen for TSendC Block
                              #statTsendcLen := #statSendBufferPos; // Buffer pos equals amount of elements in send array
                              //reset buffer pos
                              #statSendBufferPos := 0;
                              //enable Send Req
                              #statTsendcReq := TRUE;
                              //Set Watchdog
                              #statEnableTimerCommandWatchdog := TRUE;
                              //wait for send to be done
                              #statMqttCommandState := ;
                            END_IF;
                          END_IF;
                        END_REGION UNSUBSCRIBE_FROM_TOPIC

                      :
                        REGION SEND_UNSUBSCRIBE_WAIT_FOR_RESPONSE
                          //check tsend status
                          IF NOT #tempTsendcBusy AND #tempTsendcStatus =  THEN
                            IF (#statUnsubscribeTopicEncodeState = ) THEN
                              //Encoding done all sent
                              #statPaketHeaderEncodeDone := FALSE;
                            ELSE
                              // More to Encode and send
                              #statEnableTimerCommandWatchdog := FALSE;
                              #statMqttCommandState := ;
                            END_IF;
                          END_IF;
                          // Wait for timeout
                          IF #instTimerCommandWatchdog.Q THEN
                            #statEnableTimerCommandWatchdog := FALSE;
                            #statStatus := ; // Set correct status that identifies error clearly
                            #statSubfunctionStatus := ; // Status or return value of called FBs, FCs and system blocks
                            #statFBErrorState := #statFBState; // Set error state number for diagnostic
                            #statErrorAutoCleared := TRUE;
                            #statMqttCommandState := ;
                          END_IF;
                          //Check Unsubscribe ACK paket
                          CASE #tempMqttUnSubAckRcv OF
                            :  // Statement section case 1
                              ;
                            :  // Statement section case 2 to 4
                              //disable watchdog
                              #statEnableTimerCommandWatchdog := FALSE;
                              //Encoding done all sent
                              #statPaketHeaderEncodeDone := FALSE;
                              // Job done
                              #statDone := TRUE;
                              #statMqttCommandState := ;
                              // Set Status back to connected
                              #statStatus := ;
                            :
                              #statStatus := ; // Set correct status that identifies error clearly
                              #statSubfunctionStatus := ; // Status or return value of called FBs, FCs and system blocks
                              #statFBErrorState := #statFBState; // Set error state number for diagnostic
                              #statErrorAutoCleared := TRUE;
                              #statMqttCommandState := ;
                          END_CASE;
                        END_REGION SEND_UNSUBSCRIBE_WAIT_FOR_RESPONSE

                      :
                        REGION SEND_PING
                          //Set Status
                          #statStatus := ;
                          IF #tempTsendcBusy = FALSE // when tsendC is ready
                            AND #tempTsendcDone = FALSE // tsendC did not finish in this cycle
                            AND #statTsendcReq = FALSE // TsendC request was not already requested by pub ack msg
                          THEN
                            //Init
                            #statSendBufferPos := 0;
                            #statSendBuffer[#statSendBufferPos] := ;
                            #statSendBufferPos += 1;
                            //Remaining Lenght (must be 0)
                            #statSendBuffer[#statSendBufferPos] := 0;
                            #statSendBufferPos += 1;
                            #statTsendcLen := #statSendBufferPos;
                            //Start send request
                            #statTsendcReq := TRUE;
                            //Start watchdoc
                            #statEnableTimerCommandWatchdog := true;
                            //Next state
                            #statMqttCommandState := ;
                          END_IF;
                        END_REGION MQTT_COMMAND_SEND_PING

                      :
                        REGION WAIT_FOR_PING_RESP
                          //Check, if Edge of Publish comes while ping
                          IF #tempCommandInput > 0 AND NOT #statCommandInputOld THEN
                            #statCommandInputBackup := #tempCommandInput;
                            #statCommandInputOld := true;
                          END_IF;
                          //check watchdog status
                          IF #instTimerCommandWatchdog.Q THEN
                            #statEnableTimerCommandWatchdog := FALSE;
                            #statStatus := ; // Set correct status that identifies error clearly
                            #statSubfunctionStatus := ; // Status or return value of called FBs, FCs and system blocks
                            #statFBErrorState := #statFBState; // Set error state number for diagnostic
                            #statErrorAutoCleared := TRUE;
                            #statMqttCommandState := ;
                          END_IF;
                          //Check PingRsp paket
                          CASE #tempMqttPingRspRcv OF
                            :  // Statement section case 1
                              ;
                            :
                              //disable watchdog
                              #statEnableTimerCommandWatchdog := FALSE;
                              //Go to no processing
                              #statMqttCommandState := ;
                              //set Status
                              #statStatus := ;
                              IF #statCommandInputBackup <> 0 THEN
                                #statMqttCommandState := BYTE_TO_DINT(#statCommandInputBackup);
                                #statCommandInputBackup := 0;
                                #statCommandInputOld := false;
                              END_IF;
                          END_CASE;
                        END_REGION MQTT_COMMAND_PING_RESP
                      ELSE  // Statement section ELSE
                        REGION ERROR_MULTIPLE_INPUT
                          #statMqttCommandState := ; // reset back to idle
                          #statStatus := ; // Set correct status that identifies error clearly
                          #statSubfunctionStatus := ; // Status or return value of called FBs, FCs and system blocks
                          #statFBErrorState := #statFBState; // Set error state number for diagnostic
                          #statErrorAutoCleared := TRUE;
                        END_REGION ERROR_MULTIPLE_INPUT
                    END_CASE;
                  END_REGION

                  REGION CHECK_PING_TIMER
                    //If no job is running check if keepalive experied
                    IF #statMqttCommandState =
                      AND #instMqttKeepAliveTimer.Q THEN
                      //reset the timer
                      RESET_TIMER(#instMqttKeepAliveTimer);
                      //go to ping state
                      #statMqttCommandState := ;
                    END_IF;
                  END_REGION CHECK_PING_TIMER

                  //Edge detection "publish / subscribe/unsubscribe" input
                  #statPublishOld := #tempPublish;
                  #statSubscribeOld := #tempSubscribe;
                  #statUnsubscribeOld := #tempUnsubscribe;
                END_REGION CONNECTED

              ELSE   // Undefined state in state machine reached
                #statStatus := ;
                #statErrorUserCleared := TRUE;
            END_CASE;

          END_REGION MQTT_STATE_MACHINE
        END_IF;
      END_REGION FB_OPERATING_MONITOR_TCP

    :
      REGION FB_STATE_TCP_RECONNECTING
        IF #tempTsendcStatus =  THEN
          #statErrorAutoCleared := FALSE;
          // Update edge detection
          #statPublishOld := #tempPublish;
          #statSubscribeOld := #tempSubscribe;
          #statUnsubscribeOld := #tempUnsubscribe;
          //Monitor Connection
          #statFBState := ;
          // Begin MQTT Connection
          #statMqttConnectState := ;
        END_IF;
      END_REGION FB_STATE_TCP_RECONNECTING
    : // Disabling active
      REGION DISABLING FB
        //  Disabling, e.g. closing connections, etc.
        // When disabling is complete the bit #statDisablingCompleted must be set
        // When MQTT is connected, send disconnect
        IF #statMqttConnectState =  THEN
          IF #statTsendcReq = TRUE THEN
            //Interrupt any existing send jobs
            #statTsendcReq := FALSE;
          ELSE
            // INIT
            #statSendBufferPos := 0;
            //Build fixed Header
            //Message Type
            #statSendBuffer[#statSendBufferPos] := ;
            #statSendBufferPos += 1;
            //Remaining Length (must be O)
            #statSendBuffer[#statSendBufferPos] := ;
            #statSendBufferPos += 1;
            //send request
            #statTsendcLen := #statSendBufferPos;
            #statTsendcReq := TRUE;
            #statMqttConnectState := ;
          END_IF;
        ELSE
          //Disable TCP Connection
          #statTsendcReq := FALSE;
          #statTsendcEnable := FALSE;
          #statEnableTimerCommandWatchdog := TRUE;
        END_IF;
        // When TCP connection is closed
        IF #tempTsendcStatus =  THEN
          #statEnableTimerCommandWatchdog := FALSE;
          #statDisablingCompleted := TRUE;
        ELSIF #instTimerCommandWatchdog.Q THEN
          #statEnableTimerCommandWatchdog := FALSE;
          #statDisablingCompleted := TRUE;
        END_IF;
      END_REGION DISABLING FB
    ELSE // Undefined state in state machine reached
      #statStatus := ;
      #statErrorUserCleared := TRUE;
  END_CASE;
END_REGION STATE_MACHINE

REGION OUTPUTS
  // Write outputs
  IF (#statDisablingCompleted = TRUE) THEN
    // Reset outputs if disabling completed
    #statValid := FALSE;
    #statBusy := FALSE;
    #statError := FALSE;
    #statDone := FALSE;
    #statErrorUserCleared := FALSE;
    #statErrorAutoCleared := FALSE;
    #statStatus := ;
    // Reset application specific outputs
    #statRcvMsgStatus := ;
    #statRcvMsgDataLen := 0;

  ELSIF (#statErrorUserCleared = TRUE) AND (#statError = FALSE) THEN
    // Error can only be cleared by user; rising edge at enable input is needed to continue
    #statValid := FALSE;
    #statBusy := FALSE;
    #statDone := FALSE;
    #statError := TRUE;
    // Write diagnostics
    #diagnostics.status := #statStatus;
    #diagnostics.subfunctionStatus := #statSubfunctionStatus;
    #diagnostics.stateNumber := #statFBErrorState;
    // execution aborted --> set state no processing
    #statTsendcEnable := FALSE; // Terminate Connection, no reason keep it up.
    #statFBState := ;
    #statMqttConnectState := ;
    #statMqttCommandState := ;
    #statRcvMsgDecodeState := ;

  ELSIF (#statErrorAutoCleared = TRUE) AND (#statError = FALSE) THEN
    // Error can be reset by FB automatically
    #statValid := FALSE;
    #statBusy := TRUE;
    #statError := TRUE;
    #statDone := FALSE;

    // Write diagnostics
    #diagnostics.status := #statStatus;
    #diagnostics.subfunctionStatus := #statSubfunctionStatus;
    #diagnostics.stateNumber := #statFBErrorState;
    // Handling of autocleared error
    CASE #statStatus OF
        //Just signal error and reset autocleared error afterwards.
      , , ,
      , , ,
      , , :
        #statErrorAutoCleared := FALSE;

      ELSE  // Statement section ELSE
        ;
    END_CASE;

  ELSIF (#statErrorAutoCleared = FALSE) AND (#statErrorUserCleared = FALSE) AND (#statError = TRUE) THEN
    // If autocleared error is acknowledged
    #statValid := TRUE;
    #statBusy := TRUE;
    #statError := FALSE;
    #statDone := FALSE;

    //   this line  more detailed status information is used instead of "#STATUS_SUBSEQUENT_CALL"
    CASE #statStatus OF
      , :  // Reconnecting ok, start Mqtt reconnnect
        //set status
        #statStatus := ;
        //in the following status codes status stays connected.
      , , ,
      , , ,
      , :
        #statStatus := ;
      ELSE  // Statement section ELSE
        ;
    END_CASE;
  END_IF;

  // Write static values to outputs
  #valid := #statValid;
  #busy := #statBusy;
  #error := #statError;
  #status := #statStatus;
  //block sets ENO automatically:
  //ENO := TRUE;
  //Write application specific static values to outputs
  #done := #statDone;
  #receivedMsgStatus := #statRcvMsgStatus;
  #receivedMsgDataLen := #statRcvMsgDataLen;
END_REGION OUTPUTS
END_FUNCTION_BLOCK